DATA_BLOCK "S12Probe"
{ S7_Optimized_Access := 'TRUE' }
VERSION : 0.1
NON_RETAIN
   VAR
      Ready : Bool;
      Marker : DInt;
      Scans : UDInt;
   END_VAR
BEGIN
END_DATA_BLOCK
